   F[5702] := 8.785445;
   F[5703] := 8.770978;
   F[5704] := 8.709491;
   F[5705] := 8.655237;
   F[5706] := 8.74566;
   F[5707] := 8.6588545;
   F[5708] := 8.648004;
   F[5709] := 8.626302;
   F[5710] := 8.644386;
   F[5711] := 8.579283;
   F[5712] := 8.586516;
   F[5713] := 8.485243;
   F[5714] := 8.532263;
   F[5715] := 8.452691;
   F[5716] := 8.5286455;
   F[5717] := 8.492476;
   F[5718] := 8.445457;
   F[5719] := 8.39482;
   F[5720] := 8.420139;
   F[5721] := 8.387587;
   F[5722] := 8.39482;
   F[5723] := 8.351418;
   F[5724] := 8.347801;
   F[5725] := 8.318866;
   F[5726] := 8.326099;
   F[5727] := 8.224827;
   F[5728] := 8.260995;
   F[5729] := 8.217592;
   F[5730] := 8.188658;
   F[5731] := 8.192274;
   F[5732] := 8.217592;
   F[5733] := 8.098235;
   F[5734] := 8.083767;
   F[5735] := 8.0910015;
   F[5736] := 8.065682;
   F[5737] := 8.065682;
   F[5738] := 8.051215;
   F[5739] := 8.051215;
   F[5740] := 8.076533;
   F[5741] := 8.015046;
   F[5742] := 7.9716434;
   F[5743] := 7.953559;
   F[5744] := 7.9354744;
   F[5745] := 7.91739;
   F[5746] := 7.913773;
   F[5747] := 7.913773;
   F[5748] := 7.884838;
   F[5749] := 7.808883;
   F[5750] := 7.787182;
   F[5751] := 7.7907987;
   F[5752] := 7.8197336;
   F[5753] := 7.8197336;
   F[5754] := 7.761863;
   F[5755] := 7.7582464;
   F[5756] := 7.700376;
   F[5757] := 7.7148438;
   F[5758] := 7.6822915;
   F[5759] := 7.685909;
   F[5760] := 7.6461225;
   F[5761] := 7.6208043;
   F[5762] := 7.570168;
   F[5763] := 7.5882525;
   F[5764] := 7.5882525;
   F[5765] := 7.5050635;
   F[5766] := 7.562934;
   F[5767] := 7.533999;
   F[5768] := 7.526765;
   F[5769] := 7.4688945;
   F[5770] := 7.472512;
   F[5771] := 7.49783;
   F[5772] := 7.421875;
   F[5773] := 7.425492;
   F[5774] := 7.349537;
   F[5775] := 7.4037905;
   F[5776] := 7.3531537;
   F[5777] := 7.3748555;
   F[5778] := 7.306134;
   F[5779] := 7.3314524;
   F[5780] := 7.3025174;
   F[5781] := 7.313368;
   F[5782] := 7.2012444;
   F[5783] := 7.2229457;
   F[5784] := 7.295284;
   F[5785] := 7.248264;
   F[5786] := 7.172309;
   F[5787] := 7.172309;
   F[5788] := 7.1614585;
   F[5789] := 7.13614;
   F[5790] := 7.0855036;
   F[5791] := 7.0746527;
   F[5792] := 7.0891204;
   F[5793] := 7.0493345;
   F[5794] := 7.071036;
   F[5795] := 7.0167823;
   F[5796] := 6.966146;
   F[5797] := 6.9516783;
   F[5798] := 6.9516783;
   F[5799] := 6.9118924;
   F[5800] := 6.922743;
   F[5801] := 6.8684897;
   F[5802] := 6.8757234;
   F[5803] := 6.8250866;
   F[5804] := 6.8757234;
   F[5805] := 6.8684897;
   F[5806] := 6.8033853;
   F[5807] := 6.7997684;
   F[5808] := 6.781684;
   F[5809] := 6.6876445;
   F[5810] := 6.756366;
   F[5811] := 6.6948786;
   F[5812] := 6.6948786;
   F[5813] := 6.7274303;
   F[5814] := 6.6731772;
   F[5815] := 6.680411;
   F[5816] := 6.6587095;
   F[5817] := 6.6225405;
   F[5818] := 6.5863714;
   F[5819] := 6.604456;
   F[5820] := 6.575521;
   F[5821] := 6.5863714;
   F[5822] := 6.5538197;
   F[5823] := 6.5212674;
   F[5824] := 6.4742475;
   F[5825] := 6.499566;
   F[5826] := 6.4489293;
   F[5827] := 6.4344616;
   F[5828] := 6.4814816;
   F[5829] := 6.35489;
   F[5830] := 6.358507;
   F[5831] := 6.362124;
   F[5832] := 6.3368053;
   F[5833] := 6.311487;
   F[5834] := 6.358507;
   F[5835] := 6.2717013;
   F[5836] := 6.289786;
   F[5837] := 6.2572336;
   F[5838] := 6.224682;
   F[5839] := 6.213831;
   F[5840] := 6.2355323;
   F[5841] := 6.184896;
   F[5842] := 6.184896;
   F[5843] := 6.1812787;
   F[5844] := 6.09809;
   F[5845] := 6.1161747;
   F[5846] := 6.137876;
   F[5847] := 6.112558;
   F[5848] := 6.0872397;
   F[5849] := 6.0257525;
   F[5850] := 6.0293694;
   F[5851] := 6.032986;
   F[5852] := 6.101707;
   F[5853] := 5.964265;
   F[5854] := 5.9787326;
   F[5855] := 5.9497976;
   F[5856] := 5.964265;
   F[5857] := 5.910012;
   F[5858] := 5.910012;
   F[5859] := 5.862992;
   F[5860] := 5.9172454;
   F[5861] := 5.834057;
   F[5862] := 5.8268228;
   F[5863] := 5.754485;
   F[5864] := 5.8376737;
   F[5865] := 5.787037;
   F[5866] := 5.7255497;
   F[5867] := 5.0311055;
   F[5868] := 4.4958043;
   F[5869] := 3.8664641;
   F[5870] := 3.1539352;
   F[5871] := 2.6511862;
   F[5872] := 2.6692708;
   F[5873] := 2.6475694;
   F[5874] := 2.6692708;
   F[5875] := 2.7379918;
   F[5876] := 2.6620371;
   F[5877] := 2.6837385;
   F[5878] := 2.6692708;
   F[5879] := 2.6692708;
   F[5880] := 2.6114004;
   F[5881] := 2.6367188;
   F[5882] := 2.6620371;
   F[5883] := 2.5788484;
   F[5884] := 2.6367188;
   F[5885] := 2.6186342;
   F[5886] := 2.6150174;
   F[5887] := 2.6077836;
   F[5888] := 2.6077836;
   F[5889] := 2.596933;
   F[5890] := 2.589699;
   F[5891] := 2.557147;
   F[5892] := 2.589699;
   F[5893] := 2.629485;
   F[5894] := 2.5788484;
   F[5895] := 2.6041667;
   F[5896] := 2.6186342;
   F[5897] := 2.5499132;
   F[5898] := 2.5607638;
   F[5899] := 2.5282118;
   F[5900] := 2.5354457;
   F[5901] := 2.589699;
   F[5902] := 2.6041667;
   F[5903] := 2.524595;
   F[5904] := 2.5028934;
   F[5905] := 2.4739583;
   F[5906] := 2.4956598;
   F[5907] := 2.513744;
   F[5908] := 2.524595;
   F[5909] := 2.5028934;
   F[5910] := 2.524595;
   F[5911] := 2.5065105;
   F[5912] := 2.5028934;
   F[5913] := 2.513744;
   F[5914] := 2.4594908;
   F[5915] := 2.4594908;
   F[5916] := 2.419705;
   F[5917] := 2.4739583;
   F[5918] := 2.5282118;
   F[5919] := 2.4414062;
   F[5920] := 2.4269388;
   F[5921] := 2.5028934;
   F[5922] := 2.4377894;
   F[5923] := 2.4594908;
   F[5924] := 2.4414062;
   F[5925] := 2.3943865;
   F[5926] := 2.4631076;
   F[5927] := 2.5028934;
   F[5928] := 2.445023;
   F[5929] := 2.4305556;
   F[5930] := 2.4377894;

END_DATA_BLOCK
